(* CODESYS project text.library
   DefaultNamespace: KOSTAL.AF2024.Core.Text
   DocFormat: reStructuredText
   Description: Text handling
   Author: Frank Dümpelmann
   Title: KOSTAL.AF2024.Core.Text
   Version: 1.0.0.0
   Company: KOSTAL GmbH & Co.KG
   Placeholder: KOSTAL.AF2024.Core.Text

Project tree, tasks and I/O mapping:
  libraries: KOSTAL.AF2024.Core.FileLogger, 1.0.0.0 (KOSTAL GmbH & Co.KG); KOSTAL.AF2024.Core.ListOf, 1.0.0.0 (KOSTAL GmbH & Co.KG); KOSTAL.AF2024.Core.Process, 1.0.0.0 (KOSTAL GmbH & Co.KG); KOSTAL.AF2024.Core.Settings, 1.0.0.0 (KOSTAL GmbH & Co.KG); KOSTAL.AF2024.Core.StringTools, 1.0.0.0 (KOSTAL GmbH & Co.KG); KOSTAL.AF2024.Core.System, 1.0.0.0 (KOSTAL GmbH & Co.KG); Tc2_Standard, 3.3.3.0 (Beckhoff Automation GmbH); Tc2_System, 3.6.2.0 (Beckhoff Automation GmbH); Tc2_Utilities, 3.5.2.0 (Beckhoff Automation GmbH)
  Base/
    Interface/
      interface I_Text: AddVar, ClearVars, FileName, GetText, GetText_Native, LoadedLanguage, NumerOfTexts, Path, State, Valid, Vars
      interface I_Text_Owner: Ex_LoadFile, Path
    function block _FB_Base [ST]: _DELETE, FB_exit, FB_init, _fClose, _fInfo, _fOpen, _fRead, _Log, _00_idle, _10_LoadFile, _11_CreateFileBuffer, _11_FileControl, _11_FileOpen, _11_FileRead, _11_Parse, _30_ProcessFailed, _30_ProcessfPassed, _99_StepFail, _100_LoopFooter, _100_LoopHeader, _100_Origin, _100_Read, _100_StepFail, _clear, _combine, _FBmain, _mergefQFileName
  DUT/
    data type _T_textVarIndex
    data type E_Source
    data type ST_E_Text
    function block T_E_Text [ST]
  Handler/
    Base/
      function block _FB_Handler_Base [ST]: _H00_Idle, _H10_Read, AddVar, ClearVars, FBmain, GetText, GetText_Native, Reset, FileExtension, FileName, LoadedLanguage, NumerOfTexts, Path, SelectedLanguage, State, Timeout, Valid, Vars, _TextDoesNotExist
    Master/
      function block FB_Handler_Master [ST]: SelectedLanguage
    Slave/
      function block FB_Handler_Slave [ST]: linkCommonText
  Project Information/
    function F_GetCompany [ST]
    function F_GetTitle [ST]
    function F_GetVersion [ST]
  Reader/
    DUT/
      data type E_THIS_Reader
    function block FB_FileReader [ST]: AddVar, ClearVars, Ex_LoadFile, FBmain, GetText, GetText_Native, FileName, LoadedLanguage, NumerOfTexts, Path, State, Timeout, Valid, Vars
  Version/
    global variables Global_Version
  global variables GVL_CONSTANT
  global variables SOURCE
*)

// DUT/_T_textVarIndex
TYPE _T_textVarIndex : UINT(GVL_CONSTANT.VAR_MIN..GVL_CONSTANT.VAR_MAX); END_TYPE

// DUT/E_Source
{attribute 'qualified_only'}
{attribute 'strict'}
TYPE E_Source :
(
	Local 	:= 0,
	Common	:= 1
);
END_TYPE

// DUT/ST_E_Text
TYPE ST_E_Text :
	STRUCT
		Source	: E_Source:= E_Source.Local;
		Number	: UINT;
	END_STRUCT
END_TYPE

// Reader/DUT/E_THIS_Reader
{attribute 'qualified_only'}
{attribute 'strict'}
TYPE E_THIS_Reader :
(
	idle := 0,
	loadFile
	//loadLanguage
) UINT;
END_TYPE

// Version/Global_Version
{attribute 'TcGenerated'}
{attribute 'no-analysis'}
{attribute 'linkalways'}
// This function has been automatically generated from the project information.
VAR_GLOBAL CONSTANT
	{attribute 'const_non_replaced'}
	stLibVersion_KOSTAL_AF2024_Core_Text : ST_LibVersion := (iMajor := 1, iMinor := 0, iBuild := 0, iRevision := 0, nFlags := 0, sVersion := '1.0.0.0');
END_VAR

// GVL_CONSTANT
{attribute 'qualified_only'}
VAR_GLOBAL CONSTANT
	{region 'text variables'}
		VAR_IDENTIFIER	: WSTRING(1):= "#";
		VAR_MIN					: UINT:= 0;
		VAR_MAX					: UINT:= 9;
	{endregion}
END_VAR

// SOURCE
{attribute 'qualified_only'}
VAR_GLOBAL
	Common	: STRING(1):= 'C';
	Local		: STRING(1):= 'L';
END_VAR

// Base/Interface/I_Text
INTERFACE I_Text EXTENDS KOSTAL_AF2024_Core_System.I_Interface

METHOD AddVar : BOOL
VAR_INPUT
	Text	: KOSTAL_AF2024_Core_Settings.T_MaxString;
END_VAR
END_METHOD

METHOD ClearVars
VAR_INPUT
END_VAR
END_METHOD

PROPERTY FileName : KOSTAL_AF2024_Core_Settings.T_MaxString_UTF8
GET
END_GET
END_PROPERTY

METHOD GetText : KOSTAL_AF2024_Core_Settings.T_MaxString

VAR_INPUT
	Number	: ST_E_Text;
END_VAR
END_METHOD

METHOD PUBLIC GetText_Native : KOSTAL_AF2024_Core_Settings.T_MaxString

VAR_INPUT
	Number	: ST_E_Text;
END_VAR
END_METHOD

PROPERTY LoadedLanguage : KOSTAL_AF2024_Core_Settings.T_MaxString_UTF8
GET
END_GET
END_PROPERTY

PROPERTY PUBLIC NumerOfTexts : UDINT
GET
END_GET
END_PROPERTY

PROPERTY PUBLIC Path : KOSTAL_AF2024_Core_Settings.T_MaxString_UTF8	//Example:	C:\Project\Text\Common\
GET
END_GET
END_PROPERTY

PROPERTY State : KOSTAL_AF2024_Core_Process.I_T_plcState
GET
END_GET
END_PROPERTY

PROPERTY PUBLIC Valid : BOOL
GET
END_GET
END_PROPERTY

PROPERTY Vars : Kostal_AF2024_Core_StringTools.I_ListOfString
GET
END_GET
END_PROPERTY

END_INTERFACE

// Base/Interface/I_Text_Owner
INTERFACE I_Text_Owner EXTENDS I_Text

METHOD Ex_LoadFile : BOOL
VAR_INPUT
	FileName	: KOSTAL_AF2024_Core_Settings.T_MaxString_UTF8;	//full qualified filename Example: C:\Project\Text\Common.csv
END_VAR
END_METHOD

PROPERTY PUBLIC Path : KOSTAL_AF2024_Core_Settings.T_MaxString_UTF8	//Example:	C:\Project\Text\Common\
SET
END_SET
END_PROPERTY

END_INTERFACE

// Base/_FB_Base
FUNCTION_BLOCK ABSTRACT _FB_Base

VAR
	_Storage		: KOSTAL_AF2024_Core_ListOf.FB_ListOfString;
	_FileName		: KOSTAL_AF2024_Core_Settings.T_MaxString_UTF8;
	_PathName		: KOSTAL_AF2024_Core_Settings.T_MaxString_UTF8;

	_fqFileName	: KOSTAL_AF2024_Core_Settings.T_MaxString_UTF8;
	
	_Variables	: KOSTAL_AF2024_Core_ListOf.FB_ListOfString;

	_LoadedFileName	: KOSTAL_AF2024_Core_StringTools.FB_Split_UTF8;
	
	_step				: KOSTAL_AF2024_Core_process.FB_processStep_Flow;
	_State			: KOSTAL_AF2024_Core_process.T_plcState;
	
	_THIS_called		: E_THIS_Reader;
	_THIS_inProcess	: E_THIS_Reader;

	{region 'Common'}
		_FileInfo	: Tc2_Utilities.FB_EnumFindFileEntry;

		_AmsNetId	: Tc2_System.T_AmsNetID:= '';	//default local
		_ePath		: Tc2_System.E_OpenPath:= E_OpenPath.PATH_GENERIC;
	
		_FileOpen		:	Tc2_System.FB_FileOpen;
		_FileRead		: Tc2_System.FB_FileRead;
		_FileClose	: Tc2_System.FB_FileClose;
	
		_hFile		: UINT;	//UINT	> Handle to open File
	
		_FileSize		: ULINT;
		_pBuffer		: POINTER TO BYTE;
		_BufferLen	: UDINT;

	{endregion}
	
	_TimeOut		: TIME:= T#5S;

	_TempDescription	: KOSTAL_AF2024_Core_Settings.T_MaxString;
	
	_init: BOOL:= TRUE;
	
	_ILogger	: KOSTAL_AF2024_Core_FileLogger.I_Logger;
	
	_mStep	: KOSTAL_AF2024_Core_process.FB_processStep_Flow;

	{region 'file read'}
		_pReadBuffer		: POINTER TO BYTE;
		_ReadBufferLen	: UDINT;

		_readedSize			: UDINT;
		_AddressLoopHeader	: INT;
	{endregion}

END_VAR

VAR CONSTANT
	_ADDRESS_IDLE						: INT:= 0;
	_ADDRESS_LOAD_FILE			: INT:= 100;
	_ADDRESS_PROCESS_PASSED	: INT:= 300;
	_ADDRESS_PROCESS_FAILED	: INT:= 400;
	
END_VAR

METHOD PROTECTED _DELETE
VAR_INPUT
END_VAR

IF _pBuffer <> 0 THEN	__DELETE(_pBuffer);	_BufferLen:= UDINT#0;	END_IF
END_METHOD

METHOD FB_exit : BOOL
VAR_INPUT
	bInCopyCode : BOOL; // if TRUE, the exit method is called for exiting an instance that is copied afterwards (online change).
END_VAR

_clear();
_DELETE();
END_METHOD

METHOD FB_init : BOOL
VAR_INPUT
	bInitRetains : BOOL; // if TRUE, the retain variables are initialized (warm start / cold start)
	bInCopyCode : BOOL;  // if TRUE, the instance afterwards gets moved into the copy code (online change)
END_VAR

_clear();
_DELETE();
END_METHOD

METHOD PROTECTED _fClose
VAR_INPUT
	Execute		: BOOL;	//TRUE > Execution state will set to bExecute. Otherwise, no change is made to the bExecute parameter.
	Execution	: BOOL;	//Activate (TRUE) or deactivate (FALSE) then process
END_VAR

IF Execute THEN	_FileClose.bExecute:= Execution;	END_IF

_FileClose
(
	sNetId		:= _AmsNetId, 
	hFile			:= _hFile, 
	bExecute	:= , 
	tTimeout	:= _TimeOut, 
	bBusy			=> , 
	bError		=> , 
	nErrId		=> 
);

IF _FileClose.bExecute AND NOT _FileClose.bBusy THEN _hFile:= UINT#0;	END_IF
END_METHOD

METHOD PROTECTED _fInfo
VAR_INPUT
	Execute		: BOOL;	//TRUE > Execution state will set to bExecute. Otherwise, no change is made to the bExecute parameter.
	Execution	: BOOL;	//Activate (TRUE) or deactivate (FALSE) then process
	CmdType		: Tc2_Utilities.E_EnumCmdType;
END_VAR

IF Execute THEN	_FileInfo.bExecute:= Execution;	_FileInfo.eCmd:= CmdType; END_IF

_FileInfo(
	sNetId:= _AmsNetId, 
	sPathName:= _fqFileName, 
	eCmd:= , 
	bExecute:= , 
	tTimeout:= _TimeOut, 
	bBusy=> , 
	bError=> , 
	nErrID=> , 
	bEOE=> , 
	stFindFile=> );
	
//_FileInfo(bExecute:= TRUE, sPathName:= _FileName, sNetId:= _AmsNetId, eCmd:= Tc2_Utilities.E_EnumCmdType.eEnumCmd_Abort, tTimeout:= _TimeOut);

//_FileClose
//(
//	sNetId		:= _AmsNetId, 
//	hFile			:= _hFile, 
//	bExecute	:= , 
//	tTimeout	:= _TimeOut, 
//	bBusy			=> , 
//	bError		=> , 
//	nErrId		=> 
//);

//IF _FileClose.bExecute AND NOT _FileClose.bBusy THEN _hFile:= UINT#0;	END_IF
END_METHOD

METHOD PROTECTED _fOpen
VAR_INPUT
	Execute		: BOOL;	//TRUE > Execution state will set to bExecute. Otherwise, no change is made to the bExecute parameter.
	Execution	: BOOL;	//Activate (TRUE) or deactivate (FALSE) then process
END_VAR

IF Execute THEN	_FileOpen.bExecute:= Execution;	END_IF

_FileOpen
(
	sNetId		:= _AmsNetId, 
	sPathName	:= _fqFileName, 
	nMode			:= Tc2_System.FOPEN_MODEREAD OR Tc2_System.FOPEN_MODEBINARY, 
	ePath			:= _ePath, 
	bExecute	:= , 
	tTimeout	:= _TimeOut, 
	bBusy			=> , 
	bError		=> , 
	nErrId		=> , 
	hFile			=> 
);

IF _FileOpen.bExecute AND NOT _FileOpen.bBusy AND NOT _FileOpen.bError THEN _hFile:= _FileOpen.hFile;	END_IF
END_METHOD

METHOD PROTECTED _fRead
VAR_INPUT
	Execute		: BOOL;	//TRUE > Execution state will set to bExecute. Otherwise, no change is made to the bExecute parameter.
	Execution	: BOOL;	//Activate (TRUE) or deactivate (FALSE) then process
END_VAR

IF Execute THEN	_FileRead.bExecute:= Execution;	END_IF

_FileRead
(
	sNetId		:= _AmsNetId, 
	hFile			:= _hFile, 
	pReadBuff	:= _pReadBuffer, 
	cbReadLen	:= _ReadBufferLen, 
	bExecute	:= , 
	tTimeout	:= _TimeOut, 
	bBusy			=> , 
	bError		=> , 
	nErrId		=> , 
	cbRead		=> , 
	bEOF			=> 
);
END_METHOD

METHOD PROTECTED _Log
VAR_INPUT
	Text	: KOSTAL_AF2024_Core_Settings.T_MaxString;
END_VAR

IF _ILogger <> 0 THEN
	_ILogger.ID:= "TextFileReader";
	_ILogger.stepNumber:= _step.actual;
	IF  _ILogger.State.success THEN _ILogger.AddLine(Text);	END_IF
END_IF
END_METHOD

METHOD PROTECTED _00_idle

_THIS_inProcess:= E_THIS_Reader.idle;

IF _step.toggle THEN

	_fInfo(Execute:= TRUE, Execution:= FALSE, CmdType:= Tc2_Utilities.E_EnumCmdType.eEnumCmd_Abort);
	//_FileInfo(bExecute:= TRUE, sPathName:= _FileName, sNetId:= _AmsNetId, eCmd:= Tc2_Utilities.E_EnumCmdType.eEnumCmd_Abort, tTimeout:= _TimeOut);

	_fRead			(Execute:= TRUE, Execution:= FALSE);
	_fOpen			(Execute:= TRUE, Execution:= FALSE);
	_fClose			(Execute:= TRUE, Execution:= TRUE);
	_FileInfo		(bExecute:= FALSE);
END_IF

IF _FileInfo.bBusy	THEN	
	_fRead(Execute:= FALSE,	Execution:= FALSE);
ELSIF	_FileRead.bExecute	THEN	
	_fRead(Execute:= TRUE,	Execution:= FALSE);
END_IF

IF _FileRead.bBusy	THEN	
	_fRead(Execute:= FALSE,	Execution:= FALSE);
ELSIF	_FileRead.bExecute	THEN	
	_fRead(Execute:= TRUE,	Execution:= FALSE);
END_IF

IF _FileClose.bBusy THEN	
	_fClose(Execute:= FALSE,	Execution:= FALSE);
ELSIF	_FileClose.bExecute	THEN	
	_fClose(Execute:= TRUE,	Execution:= FALSE);
END_IF

IF _FileOpen.bBusy	THEN	
	_fOpen(Execute:= FALSE,	Execution:= FALSE);
ELSIF	_FileOpen.bExecute	THEN	
	_fOpen(Execute:= TRUE,	Execution:= FALSE);
END_IF

_State.clear();

IF _FileOpen.bBusy 			THEN	
	_State.busy := TRUE;	
	_State.description:= "_fCommonOpen is busy. Please wait ...";
ELSIF _FileRead.bBusy	THEN	
	_State.busy := TRUE;	
	_State.description:= "_fCommonGetString is busy. Please wait ...";
ELSIF _FileClose.bBusy 			THEN	
	_State.busy := TRUE;	
	_State.description:= "_fCommonClose is busy. Please wait ...";

ELSIF _THIS_called = E_THIS_Reader.loadFile 		THEN	
	_THIS_inProcess:= E_THIS_Reader.loadFile;	
	_step.set(_ADDRESS_LOAD_FILE);

ELSE
	_State.ready:= TRUE;
END_IF
END_METHOD

METHOD PROTECTED _10_LoadFile

VAR
	_result: KOSTAL_AF2024_Core_Settings.T_MaxString;
END_VAR

_THIS_inProcess:= E_THIS_Reader.loadFile;

_State.clear();
_State.busy := TRUE;

IF _step.toggle THEN	
	_DELETE();	
	_Storage.clear();
	_FileSize:= ULINT#0;	
	_LoadedFileName.Clear();
END_IF


IF NOT _mergefQFileName(_result) THEN	_30_ProcessFailed(_result);
ELSE																	_step.INC();	
END_IF
END_METHOD

METHOD PROTECTED _11_CreateFileBuffer


IF _step.toggle THEN	
	_BufferLen:= ULINT_TO_UDINT(_FileSize);
	_pBuffer:= __NEW(BYTE, _BufferLen);	
END_IF

_State.clear();
_State.busy := TRUE;

IF _pBuffer = 0 THEN	_30_ProcessFailed("Not possible to create file buffer");
ELSE									_step.INC();	
END_IF
END_METHOD

METHOD PROTECTED _11_FileControl

IF _step.toggle THEN
	_fInfo(Execute:= TRUE, Execution:= TRUE, CmdType:= Tc2_Utilities.E_EnumCmdType.eEnumCmd_First);
	//_FileInfo(bExecute:= TRUE, sPathName:= _FileName, sNetId:= _AmsNetId, eCmd:= Tc2_Utilities.E_EnumCmdType.eEnumCmd_First, tTimeout:= _TimeOut);
END_IF

_State.clear();
_State.busy := TRUE;

_fInfo(Execute:= TRUE, Execution:= FALSE, CmdType:= Tc2_Utilities.E_EnumCmdType.eEnumCmd_First);
//_FileInfo(bExecute:= FALSE);

IF _FileInfo.bBusy THEN	

	_State.description:= "get common fileinfo is not finished... please wait";

ELSIF _FileInfo.bError	THEN

	_30_ProcessFailed("common file not able to read - retries overflow");
	
ELSE

	_FileSize:= Tc2_Utilities.ULARGE_TO_ULINT(_FileInfo.stFindFile.fileSize);

	IF 		_FileInfo.stFindFile.sFileName = ''	THEN	_30_ProcessFailed("File does not exist");
	ELSIF _FileSize = ULINT#0									THEN	_30_ProcessfPassed("File is empty");
	ELSE																						_step.INC();
	END_IF

END_IF
END_METHOD

METHOD PROTECTED _11_FileOpen

IF _step.toggle THEN
	_fOpen(TRUE, FALSE);
	_fOpen(TRUE, TRUE);
END_IF

_State.clear();
_State.busy := TRUE;

_fOpen(FALSE, FALSE);

IF _FileOpen.bBusy THEN	

	_State.description:= "open file is not finished... please wait";

ELSIF _FileOpen.bError	THEN

	_fOpen(TRUE, FALSE);
	_30_ProcessFailed(Tc2_Standard.WCONCAT("file not able to open - retries overflow; ErrID:", UDINT_TO_WSTRING(_FileOpen.nErrId)));
	
ELSE
	
	_hFile:= _FileOpen.hFile;
	
	_step.INC();

END_IF
END_METHOD

METHOD PROTECTED _11_FileRead

IF _step.toggle THEN
	_mStep.init();
END_IF


_mStep.Header();

IF _mStep.isActive(0) THEN	_100_Origin();			END_IF
IF _mStep.isActive(1) THEN	_100_LoopHeader();	END_IF
IF _mStep.isActive(2) THEN	_100_Read();				END_IF
IF _mStep.isActive(3) THEN	_100_LoopFooter();	END_IF


IF _mStep.NotFound()	THEN	_100_StepFail();	END_IF


(*
IF _step.toggle THEN
	_RetryCounter:= 0;
	_fRead(TRUE, FALSE);
	_fRead(TRUE, TRUE);
END_IF

_Status.clear();
_Status.setUnique_busy();

_fRead(TRUE, FALSE);

IF _FileRead.bBusy THEN	

	_Status.description:= 'read file is not finished... please wait';

ELSIF _FileRead.bError	THEN

	IF _RetryCounter >= _Retries	THEN
	
		_30_ProcessFailed(Tc2_Standard.CONCAT('file not able to read - retries overflow; ErrID:', UDINT_TO_STRING(_FileRead.nErrId)));
	
	ELSE
	
		_RetryCounter:= _RetryCounter + 1;

		_Status.description:= Tc2_Standard.CONCAT('common file not able to read - tryagain; ErrID:', UDINT_TO_STRING(_FileRead.nErrId));
		_Log(_Status.description);
		
		_fRead(TRUE, FALSE);
		_fRead(TRUE, TRUE);

	END_IF

ELSIF _FileRead.cbRead <> _FileSize	THEN

	IF _RetryCounter >= _Retries	THEN
	
		_30_ProcessFailed(Tc2_Standard.CONCAT('file not able to read completely - retries overflow; ErrID:', UDINT_TO_STRING(_FileRead.nErrId)));
	
	ELSE
	
		_RetryCounter:= _RetryCounter + 1;

		_Status.description:= Tc2_Standard.CONCAT('common file not able to read completely - tryagain; ErrID:', UDINT_TO_STRING(_FileRead.nErrId));
		_Log(_Status.description);
		
		_fRead(TRUE, FALSE);
		_fRead(TRUE, TRUE);

	END_IF

ELSE
	
	_step.INC();

END_IF

*)
END_METHOD

METHOD PROTECTED _11_Parse

VAR
	_udi: UDINT;

	_pWs1	: POINTER TO WSTRING(1);
	_ws1	: WSTRING(1);
	_wTemp	: KOSTAL_AF2024_Core_Settings.T_MaxString;
	_pWord: POINTER TO WORD;
	_Swap: BOOL;
	_StartCount: UDINT;
END_VAR

IF _step.toggle THEN	;	END_IF	

_State.clear();
_State.busy := TRUE;

_wTemp:= "";

{region 'LE/BE Endian detection'}
	//select Big or little endian (TC works with little endian)
	_pWord:= _pBuffer;
	
	IF _pWord^ = KOSTAL_AF2024_Core_Settings.GVL_CONSTANT.UNICODE_BigEndian THEN
		_Swap:= TRUE;
		_StartCount:= 2;
	ELSIF _pWord^ = KOSTAL_AF2024_Core_Settings.GVL_CONSTANT.UNICODE_LittleEndian THEN
		_Swap:= FALSE;
		_StartCount:= 2;
	ELSE
		_Swap:= FALSE;
		_StartCount:= 2;
	END_IF
{endregion}

FOR _udi:= _StartCount TO _BufferLen - 2 BY 2 DO

 	_pWord:= _pBuffer + _udi;

	//swap to little endian
	IF _Swap THEN	_pWord^:= Tc2_Utilities.BE16_TO_HOST(_pWord^);	END_IF

	_pWs1:= _pWord;
	_ws1:= _pWs1^; 

	IF _ws1 = "$R" THEN
		_Storage.addLine(_wTemp);
		_wTemp:= "";
	ELSIF _ws1 = "$N" THEN	;	//do nothing
	//ELSIF _ws1 = "" 	THEN	;	//do nothing
	ELSE	_wTemp:= Tc2_Standard.WCONCAT(_wTemp, _ws1);
	END_IF

END_FOR

_step.INC();
END_METHOD

METHOD PROTECTED _30_ProcessFailed
VAR_INPUT
	Description	: KOSTAL_AF2024_Core_Settings.T_MaxString;
END_VAR

IF _step.actual <> _ADDRESS_PROCESS_FAILED THEN _TempDescription:= Description;	_step.set(_ADDRESS_PROCESS_FAILED);	RETURN;	END_IF

IF _step.toggle THEN
	_log(_TempDescription);
END_IF

_State.clear();
_State.fail				:= TRUE;
_State.description	:= _TempDescription;
_State.finish			:= TRUE;
END_METHOD

METHOD PROTECTED _30_ProcessfPassed
VAR_INPUT
	Description	: KOSTAL_AF2024_Core_Settings.T_MaxString;
END_VAR

IF _step.actual <> _ADDRESS_PROCESS_PASSED THEN _TempDescription:= Description;	_step.set(_ADDRESS_PROCESS_PASSED);	RETURN;	END_IF

IF _step.toggle THEN
	_LoadedFileName.Split_Delimiter(_FileName, '.');
	_log(_TempDescription);
END_IF

_State.clear();
_State.pass				:= TRUE;
_State.description	:= _TempDescription;
_State.finish			:= TRUE;
END_METHOD

METHOD PROTECTED _99_StepFail
VAR_INPUT
END_VAR

_State.clear();
_State.fail:= TRUE;
_State.description:= Tc2_Standard.WCONCAT("STEP does not exist: ", INT_TO_WSTRING(_step.actual));

IF _step.toggle THEN	_Log(_State.description);	END_IF
END_METHOD

METHOD PROTECTED _100_LoopFooter
VAR_INPUT
END_VAR

IF _mStep.toggle	THEN	;	END_IF

//finished
IF (_readedSize >= _BufferLen) OR _FileRead.bEOF	THEN
	
	_step.INC();

ELSE

	_mStep.set(_AddressLoopHeader);

END_IF
END_METHOD

METHOD PROTECTED _100_LoopHeader
VAR_INPUT
END_VAR

IF _mStep.toggle	THEN	;	END_IF

_AddressLoopHeader:= _mStep.actual;

_mStep.INC();
END_METHOD

METHOD PROTECTED _100_Origin
VAR_INPUT
END_VAR

IF _mStep.toggle THEN
	_readedSize			:= UDINT#0;
	_pReadBuffer		:= _pBuffer;
	_ReadBufferLen	:= _BufferLen;
END_IF

_mStep.INC();
END_METHOD

METHOD PROTECTED _100_Read
VAR_INPUT
END_VAR

IF _mStep.toggle THEN
	_fRead(TRUE, FALSE);
	_fRead(TRUE, TRUE);
END_IF

_fRead(FALSE, TRUE);

IF _FileRead.bBusy THEN	

	_State.description:= "read file is not finished... please wait";

ELSIF _FileRead.bError	THEN

	_30_ProcessFailed(Tc2_Standard.WCONCAT("file not able to read; ErrID:", UDINT_TO_WSTRING(_FileRead.nErrId)));

ELSE
	
	_readedSize:= _readedSize + _FileRead.cbRead;
	_pReadBuffer:= _pBuffer + _readedSize;
	_ReadBufferLen:= _BufferLen - _readedSize;
	
	_mStep.INC();

END_IF
END_METHOD

METHOD PROTECTED _100_StepFail
VAR_INPUT
END_VAR

_State.clear();
_State.fail:= TRUE;
_State.description:= Tc2_Standard.WCONCAT(" _mStep(FileRead) _Step does not exist: ", INT_TO_WSTRING(_mStep.actual));

IF _mStep.toggle THEN	_Log(_State.description);	END_IF
END_METHOD

METHOD PROTECTED _clear
VAR_INPUT
END_VAR

_LoadedFileName.Clear();
_Storage.clear();
_Variables.clear();
END_METHOD

(*
Description
===========
| Protected method - to be used in derived function blocks only!
| Replace all variables in text by strings from variable table
| Parameters:
| 	text: STRING(255): Text to replace variables in
| Returns: String(255) with replaced variables

*)

METHOD PROTECTED _combine : KOSTAL_AF2024_Core_Settings.T_MaxString
VAR_INPUT
	Text	: KOSTAL_AF2024_Core_Settings.T_MaxString;
END_VAR

VAR
	_text			: KOSTAL_AF2024_Core_Settings.T_MaxString;
	_var			: KOSTAL_AF2024_Core_Settings.T_MaxString;
	_i				: INT;
	_varIndex	: _T_textVarIndex;
	_reload		: BOOL;
END_VAR

_text:= Text;

IF _Variables.NumberOfLines = 0			 															THEN	;	//no Variables available
ELSIF Tc2_Standard.WFIND(_text, GVL_CONSTANT.VAR_IDENTIFIER) = 0	THEN	;	//no Variables in Text available
	
ELSE

	_reload:= FALSE;
	
	_i:= 1;
	
	//search until the second last position
	REPEAT
	
		
		//get Position of Variable identifier
		IF Tc2_Standard.WMID(_text, 1, _i) = GVL_CONSTANT.VAR_IDENTIFIER THEN
	
			//identifier found
			_varIndex:= WSTRING_TO_UINT(Tc2_Standard.WMID(_text, 1, _i + 1)); 
	
			IF _varIndex > 0 OR (Tc2_Standard.WMID(_text, 1, _i + 1) = "0") THEN
				_var:= _Variables.line_GET(_varIndex + 1);
				_text:= Tc2_Standard.WREPLACE(_text, _var, 2, _i);
				_reload:= TRUE;
			END_IF
	
		END_IF

		//decrement counter (-1) if Identifier was found  
		IF _reload THEN	_reload:= FALSE;
		ELSE						_i:=_i + 1;		
		END_IF


	UNTIL _i >= Tc2_Standard.WLEN(_text)
	END_REPEAT
	
END_IF

_combine:= _text;
END_METHOD

METHOD PROTECTED _FBmain
VAR_INPUT
END_VAR

IF (_THIS_called <> _THIS_inProcess) AND (_step.actual <> _ADDRESS_IDLE) OR _init THEN	_step.init();	END_IF

_step.Header();


IF _step.isActive(_ADDRESS_IDLE)	THEN _00_idle();	END_IF


IF _step.isActive(_ADDRESS_LOAD_FILE)			THEN _10_LoadFile();					END_IF
IF _step.isActive(_ADDRESS_LOAD_FILE + 1)	THEN _11_FileControl();				END_IF
IF _step.isActive(_ADDRESS_LOAD_FILE + 2)	THEN _11_CreateFileBuffer();	END_IF
IF _step.isActive(_ADDRESS_LOAD_FILE + 3)	THEN _11_FileOpen();					END_IF
IF _step.isActive(_ADDRESS_LOAD_FILE + 4)	THEN _11_FileRead();					END_IF
IF _step.isActive(_ADDRESS_LOAD_FILE + 5)	THEN _11_Parse();							END_IF
IF _step.isActive(_ADDRESS_LOAD_FILE + 6)	THEN _30_ProcessfPassed("File loaded successfully");	END_IF

IF _step.isActive(_ADDRESS_PROCESS_PASSED)	THEN _30_ProcessfPassed("");	END_IF

IF _step.isActive(_ADDRESS_PROCESS_FAILED)	THEN _30_ProcessFailed("");	END_IF


IF _step.NotFound()	THEN	_99_StepFail();	END_IF



_init:= FALSE;
END_METHOD

METHOD PROTECTED _mergefQFileName : BOOL
VAR_INPUT
	Result	: REFERENCE TO KOSTAL_AF2024_Core_Settings.T_MaxString;
END_VAR

IF _PathName = '' THEN	
	IF __ISVALIDREF(Result)	THEN Result:= "Pathname is empty";	END_IF
	RETURN;	
END_IF

IF _FileName = '' THEN	
	IF __ISVALIDREF(Result)	THEN Result:= "Filename is empty";	END_IF
	RETURN;	
END_IF

IF Tc2_Standard.RIGHT(_PathName, 1) <> '\' THEN	
	_PathName:= Tc2_Standard.CONCAT(_PathName, '\');
END_IF

IF Tc2_Standard.LEFT(_FileName, 1) = '\' THEN	
	_FileName:= Tc2_Standard.RIGHT(_FileName, Tc2_Standard.LEN(_FileName) - 1);
END_IF

_fqFileName:= Tc2_Standard.CONCAT(_PathName, _FileName);

IF __ISVALIDREF(Result)	THEN Result:= "successful";	END_IF

_mergefQFileName:= TRUE;
END_METHOD

END_FUNCTION_BLOCK

// DUT/T_E_Text
FUNCTION_BLOCK PUBLIC T_E_Text

END_FUNCTION_BLOCK

// Handler/Base/_FB_Handler_Base
FUNCTION_BLOCK _FB_Handler_Base EXTENDS _FB_Base IMPLEMENTS I_Text
VAR_STAT
	_SELECTED_LANGUAGE	: KOSTAL_AF2024_Core_Settings.T_MaxString_UTF8;
END_VAR

VAR
	_H_Step	: KOSTAL_AF2024_Core_process.FB_processStep_Flow;
	_Reset	: BOOL;
	_FileExtension	: KOSTAL_AF2024_Core_Settings.T_MaxString_UTF8:= '.txt';
	_loadLanguage: KOSTAL_AF2024_Core_Settings.T_MaxString_UTF8;

	{region 'CommonText'}
		_CommonText	: I_Text;
	{endregion}
END_VAR

VAR CONSTANT
	_H_ADDRESS_IDLE	: INT:= 0;
END_VAR

METHOD PROTECTED _H00_Idle

var
	_c	: Kostal_AF2024_Core_StringTools.FB_Concat_UTF8;
END_VAR

IF _Reset THEN _Reset:= FALSE;
	
ELSIF _THIS_inProcess <> E_THIS_Reader.idle	THEN	;

ELSIF NOT _State.ready	THEN	;
	
ELSIF (_SELECTED_LANGUAGE = '') THEN

_State.clear();
_State.description:= "No language is requested"; 

ELSIF (_SELECTED_LANGUAGE <> '') AND (_SELECTED_LANGUAGE <> _LoadedFileName.Results.line_GET(1)) THEN

	_loadLanguage:= _SELECTED_LANGUAGE;
	
	_c.Clear();
	_c.addContent(_loadLanguage);
	_c.addContent(_FileExtension);
	
	_FileName:= _c.getResult();
	
	_c.Clear();
	
	_H_Step.INC();

END_IF
END_METHOD

METHOD PROTECTED _H10_Read

_THIS_called:= E_THIS_Reader.loadFile;


_THIS_called:= E_THIS_Reader.loadFile;

_FBmain();

IF NOT _State.finish 										THEN	;
ELSIF _State.pass 												THEN	_H_Step.set(_H_ADDRESS_IDLE);	
ELSIF _loadLanguage <> _SELECTED_LANGUAGE	THEN	_H_Step.set(_H_ADDRESS_IDLE);
END_IF
END_METHOD

METHOD AddVar : BOOL
VAR_INPUT
	Text	: KOSTAL_AF2024_Core_Settings.T_MaxString;
END_VAR

AddVar:= _Variables.addLine(Text);
END_METHOD

METHOD ClearVars

_Variables.clear();
END_METHOD

METHOD PUBLIC FBmain
VAR_INPUT
END_VAR

IF _init OR _Reset THEN	_H_Step.init();	_Reset:= FALSE;	END_IF

_H_Step.Header();

IF _H_Step.isActive(0) THEN	_H00_Idle();	END_IF
IF _H_Step.isActive(1) THEN	_H10_Read();	END_IF




 
 


IF _THIS_called = E_THIS_Reader.idle THEN
	_FBmain();
END_IF

_THIS_called:= E_THIS_Reader.idle;
END_METHOD

METHOD GetText : KOSTAL_AF2024_Core_Settings.T_MaxString

VAR_INPUT
	Number	: ST_E_Text;
END_VAR

VAR
	_Native: KOSTAL_AF2024_Core_Settings.T_MaxString;
END_VAR


IF Number.Number = 0 THEN GetText:= _TextDoesNotExist(Number);	RETURN;	END_IF

IF Number.Source = E_Source.Common THEN	//common Text
	
	IF _CommonText = 0	THEN GetText:= "Common Text is not linked";	RETURN;	END_IF

	Number.Source:= E_Source.Local;
	_Native	:= _CommonText.GetText_Native(Number);

	GetText:= SUPER^._combine(_Native);

ELSE	//local Text

	GetText:= _combine(_Storage.line_GET(Number.Number));
	
END_IF

IF GetText = "" THEN	GetText:= _TextDoesNotExist(Number);	END_IF
END_METHOD

METHOD PUBLIC GetText_Native : KOSTAL_AF2024_Core_Settings.T_MaxString

VAR_INPUT
	Number	: ST_E_Text;
END_VAR


IF Number.Number = 0 THEN GetText_Native:= _TextDoesNotExist(Number);	RETURN;	END_IF

IF Number.Source = E_Source.Common THEN	//common Text
	
	IF _CommonText = 0	THEN GetText_Native:= "Common Text is not linked";	RETURN;	END_IF

	Number.Source:= E_Source.Local;
	GetText_Native	:= _CommonText.GetText_Native(Number);

ELSE

		GetText_Native:= _Storage.line_GET(Number.Number);

END_IF
	
IF GetText_Native = "" THEN	GetText_Native:= _TextDoesNotExist(Number);	END_IF
END_METHOD

METHOD PUBLIC Reset
VAR_INPUT
END_VAR

_Reset:= TRUE;
END_METHOD

PROPERTY PUBLIC FileExtension : KOSTAL_AF2024_Core_Settings.T_MaxString_UTF8
GET
END_GET
SET
END_SET
END_PROPERTY

PROPERTY FileName : KOSTAL_AF2024_Core_Settings.T_MaxString_UTF8
GET

FileName:= _FileName;
END_GET
END_PROPERTY

PROPERTY LoadedLanguage : KOSTAL_AF2024_Core_Settings.T_MaxString_UTF8
GET

LoadedLanguage:= _LoadedFileName.Results.line_GET(1); //WSTRING_TO_STRING(_Storage.line_GET(KOSTAL_AF2024_Core_Settings.GVL_CONSTANT.TEXT_LINE_LANGUAGE_NAME));
END_GET
END_PROPERTY

PROPERTY PUBLIC NumerOfTexts : UDINT
GET

NumerOfTexts:= _Storage.NumberOfLines;
END_GET
END_PROPERTY

PROPERTY PUBLIC Path : KOSTAL_AF2024_Core_Settings.T_MaxString_UTF8	//Example:	C:\Project\Text\Common\
GET

Path:= _PathName;
END_GET
SET

_PathName:= Path;
END_SET
END_PROPERTY

PROPERTY SelectedLanguage : KOSTAL_AF2024_Core_Settings.T_MaxString_UTF8
GET

SelectedLanguage:= _SELECTED_LANGUAGE;
END_GET
END_PROPERTY

PROPERTY State : KOSTAL_AF2024_Core_Process.I_T_plcState
GET

State:= _State;
END_GET
END_PROPERTY

PROPERTY PUBLIC Timeout : TIME
GET

Timeout:= _TimeOut;
END_GET
SET

IF Timeout < T#5S THEN	_TimeOut:= T#5S;	
ELSE										_TimeOut:= Timeout;
END_IF
END_SET
END_PROPERTY

PROPERTY PUBLIC Valid : BOOL
GET

Valid:= 		_State.ready 
	AND_THEN (_loadLanguage <> '') 
	AND_THEN (_Storage.NumberOfLines <> 0) 
	AND_THEN (_THIS_called = E_THIS_Reader.idle) 
	AND_THEN NOT _Reset;
END_GET
END_PROPERTY

PROPERTY Vars : Kostal_AF2024_Core_StringTools.I_ListOfString
GET

Vars:= _Variables;
END_GET
END_PROPERTY

METHOD PROTECTED _TextDoesNotExist : KOSTAL_AF2024_Core_Settings.T_MaxString
VAR_INPUT
	Number	: ST_E_Text;
END_VAR

VAR
	_c: Kostal_AF2024_Core_StringTools.FB_Concat;
END_VAR

_c.Clear();
_c.addContent("#Text Number >");
_c.addContent(UINT_TO_WSTRING(Number.Number));

IF Number.Source = E_Source.Common THEN
	_c.addContent("< from Common Text does not exist or is empty#");
ELSE
	_c.addContent("< from Local Text does not exist or is empty#");
END_IF

_TextDoesNotExist := _c.getResult();
END_METHOD

END_FUNCTION_BLOCK

// Handler/Master/FB_Handler_Master
FUNCTION_BLOCK FB_Handler_Master EXTENDS _FB_Handler_Base

PROPERTY SelectedLanguage : KOSTAL_AF2024_Core_Settings.T_MaxString_UTF8
SET

_SELECTED_LANGUAGE:= SelectedLanguage;
END_SET
END_PROPERTY

END_FUNCTION_BLOCK

// Handler/Slave/FB_Handler_Slave
FUNCTION_BLOCK FB_Handler_Slave EXTENDS _FB_Handler_Base

METHOD PUBLIC linkCommonText
VAR_INPUT
	Common	: I_Text;
END_VAR

_CommonText:= Common;
END_METHOD

END_FUNCTION_BLOCK

// Project Information/F_GetCompany
// This function has been automatically generated from the project information.
{attribute 'signature_flag' := '1073741824'}
{attribute 'TcGenerated'}
{attribute 'no-analysis'}
FUNCTION F_GetCompany : WSTRING
VAR_INPUT
	
END_VAR

F_GetCompany := "KOSTAL GmbH & Co.KG";

END_FUNCTION

// Project Information/F_GetTitle
// This function has been automatically generated from the project information.
{attribute 'signature_flag' := '1073741824'}
{attribute 'TcGenerated'}
{attribute 'no-analysis'}
FUNCTION F_GetTitle : WSTRING
VAR_INPUT
	
END_VAR

F_GetTitle := "KOSTAL.AF2024.Core.Text";

END_FUNCTION

// Project Information/F_GetVersion
// This function has been automatically generated from the project information.
{attribute 'signature_flag' := '1073741824'}
{attribute 'TcGenerated'}
{attribute 'no-analysis'}
FUNCTION F_GetVersion : ST_LibVersion
VAR_INPUT
	
END_VAR

F_GetVersion.iMajor := 1;
F_GetVersion.iMinor := 0;
F_GetVersion.iBuild := 0;
F_GetVersion.iRevision := 0;
F_GetVersion.sVersion := '1.0.0.0';
F_GetVersion.nFlags := 0;

END_FUNCTION

// Reader/FB_FileReader
FUNCTION_BLOCK FB_FileReader EXTENDS _FB_Base IMPLEMENTS I_Text, I_Text_Owner

METHOD AddVar : BOOL
VAR_INPUT
	Text	: KOSTAL_AF2024_Core_Settings.T_MaxString;
END_VAR

AddVar:= _Variables.addLine(Text);
END_METHOD

METHOD ClearVars

_Variables.clear();
END_METHOD

METHOD Ex_LoadFile : BOOL
VAR_INPUT
	FileName	: KOSTAL_AF2024_Core_Settings.T_MaxString_UTF8;	//only file nameExample: English.txt
END_VAR
IF _THIS_called = E_THIS_Reader.idle THEN

	_FileName:= FileName;

	_THIS_called:= E_THIS_Reader.loadFile;

	_FBmain();

	Ex_LoadFile:= _THIS_called = _THIS_inProcess;

END_IF
END_METHOD

METHOD PUBLIC FBmain
VAR_INPUT
END_VAR

IF _THIS_called = E_THIS_Reader.idle THEN
	_FBmain();
END_IF

_THIS_called:= E_THIS_Reader.idle;
END_METHOD

METHOD PUBLIC GetText : KOSTAL_AF2024_Core_Settings.T_MaxString

VAR_INPUT
	Number	: ST_E_Text;
END_VAR

GetText:= "";

IF Number.Number = 0 THEN RETURN;	END_IF

GetText:= _combine(_Storage.line_GET(Number.Number));
END_METHOD

METHOD PUBLIC GetText_Native : KOSTAL_AF2024_Core_Settings.T_MaxString

VAR_INPUT
	Number	: ST_E_Text;
END_VAR

GetText_Native:= "";

IF Number.Number = 0 THEN RETURN;	END_IF

GetText_Native:= _Storage.line_GET(Number.Number);
END_METHOD

PROPERTY FileName : KOSTAL_AF2024_Core_Settings.T_MaxString_UTF8
GET

FileName:= _FileName;
END_GET
END_PROPERTY

PROPERTY LoadedLanguage : KOSTAL_AF2024_Core_Settings.T_MaxString_UTF8
GET

LoadedLanguage:= _LoadedFileName.Results.line_GET(1);
END_GET
END_PROPERTY

PROPERTY PUBLIC NumerOfTexts : UDINT
GET

NumerOfTexts:= _Storage.NumberOfLines;
END_GET
END_PROPERTY

PROPERTY PUBLIC Path : KOSTAL_AF2024_Core_Settings.T_MaxString_UTF8	//Example:	C:\Project\Text\Common\
GET

Path:= _PathName;
END_GET
SET

_PathName:= Path;
END_SET
END_PROPERTY

PROPERTY State : KOSTAL_AF2024_Core_process.I_T_plcState
GET

State:= _State;
END_GET
END_PROPERTY

PROPERTY PUBLIC Timeout : TIME
GET

Timeout:= _TimeOut;
END_GET
SET

IF Timeout < T#5S THEN	_TimeOut:= T#5S;	
ELSE										_TimeOut:= Timeout;
END_IF
END_SET
END_PROPERTY

PROPERTY PUBLIC Valid : BOOL
GET

Valid:= 		_State.ready 
	AND_THEN (LoadedLanguage <> '') 
	AND_THEN (_Storage.NumberOfLines <> 0) 
	AND_THEN (_THIS_called = E_THIS_Reader.idle);
END_GET
END_PROPERTY

PROPERTY Vars : Kostal_AF2024_Core_StringTools.I_ListOfString
GET

Vars:= _Variables;
END_GET
END_PROPERTY

END_FUNCTION_BLOCK
